(* ================================================================= *)
(*  FB_1030_SafetyManager                                             *)
(*  全机安全管理块: 安全回路状态 + 两次复位 + 启动许可 + 门锁开门流程   *)
(*  版本: V1.0.0  日期: 2026-10-22                                    *)
(*  来源: SysLib/safety/                                              *)
(*  依据: 电气自动化安全规范 V1.0 第 0/2/3/4/5/8/9/12 节               *)
(*        安全FB设计草案_20261022 (用户 10-22 定: 合成一块)            *)
(*  依赖: FB_TON V3.0.0 (真实毫秒), FB_R_TRIG                          *)
(*                                                                    *)
(*  它管什么:                                                         *)
(*    - 只读安全器件报给 PLC 的状态点, 算出"能不能动""复位采不采纳"    *)
(*      "能不能开门", 交给各工位块使用. 全机只调用一次.                *)
(*  它不管什么:                                                       *)
(*    - 不控制安全回路 (回路靠安全继电器硬件切断, 规范 0.1)            *)
(*    - 不决定电磁阀急停后清零还是保持 (工位块按 IO 表, 规范 2.3)       *)
(*    - 不决定断点续跑还是重新初始化 (工位块按项目需求, 规范 2.5)       *)
(*    - 不做光栅屏蔽 (规范 5.3), 不做按钮卡住判断 (规范 3.5)           *)
(*                                                                    *)
(*  状态 q_iState:                                                    *)
(*    0 安全回路断开   1 等满 10 s   2 等运行复位   3 等启动   4 运行许可 *)
(*                                                                    *)
(*  两次复位 (规范 3.1~3.6, 10 s 从第一次按复位起算, 用户 10-21 定):  *)
(*    第一次: 安全继电器自行复位, PLC 只记时刻 (门锁好、总线在线才记)  *)
(*    第二次: 继电器反馈正常 且 距第一次 >= 10 s 才采纳 -> 运行复位脉冲 *)
(*    之后按启动 -> 启动脉冲 + 运行许可. 复位/启动都只认上升沿.         *)
(*                                                                    *)
(*  报警字 q_dwAlarm:                                                 *)
(*    bit0~7   第 1~8 个急停被按下 (实时)                              *)
(*    bit8~15  第 1~8 扇门没关好/没锁 (实时)                           *)
(*    bit16~23 第 1~8 道光栅被遮挡 (实时)                              *)
(*    bit24~27 第 1~4 个安全继电器反馈 = 故障 (实时)                    *)
(*    bit28    总线断线 (实时)                                         *)
(*    bit29    复位被拒: 安全回路未恢复/门没锁/总线断 (保持到下次采纳)  *)
(*    bit30    复位过早: 距第一次不足 10 s (保持到下次采纳)             *)
(*    bit31    门锁回失败: 撤销解锁后 1 s 内门锁点没回来 (保持到锁好)   *)
(*                                                                    *)
(*  安全区: 改本块等于改安全区, 先仿真再由用户签字 (规范 0.5)         *)
(* ================================================================= *)

FUNCTION_BLOCK FB_1030_SafetyManager

VAR_INPUT
    i_arrSafetyFault : ARRAY[0..3] OF BOOL;  // 安全继电器 41-42 常闭辅助点, 1 = 安全回路故障; 未用的填 FALSE (规范 8.1, 判断的唯一依据)
    i_arrEStopOk     : ARRAY[0..7] OF BOOL;  // 急停按钮第三组触点, 1 = 正常; 未用的填 TRUE (规范 2.2, 只报警定位)
    i_arrCurtainOk   : ARRAY[0..7] OF BOOL;  // 光栅进 PLC 的状态点, 1 = 未遮挡; 未用的填 TRUE (规范 5.1, 只报警定位)
    i_arrDoorClosed  : ARRAY[0..7] OF BOOL;  // 门锁进 PLC 的那组触点, 1 = 门关好且已锁; 未用的填 TRUE (规范 4.1, 4.4)
    i_bFieldbusOk    : BOOL;                 // 远程 IO/总线伺服全部在线 (项目汇总后接入, 规范 8.3)
    i_bResetBtn      : BOOL;                 // 复位按钮进 PLC 的那组触点 (规范 3.1)
    i_bStartBtn      : BOOL;                 // 启动按钮 (规范 3.6)
    i_bAutoMode      : BOOL;                 // 设备在自动 (全机一个, 自动时申请开门不响应)
    i_bMotionStopped : BOOL;                 // 伺服零速 + 所有动作完全停止 (全机一个, 项目汇总后接入)
    i_arrDoorReqBtn  : ARRAY[0..7] OF BOOL;  // 每扇门的申请开门按钮; 未用的填 FALSE
END_VAR

VAR_OUTPUT
    q_bSafeToRun     : BOOL;                 // 1 = 可以动; 各工位块的运动输出都要和它"与" (规范 0.1)
    q_bStopNow       : BOOL;                 // 1 = 安全条件现在丢了 (继电器故障/门没锁/总线断), 同一扫描生效 (规范 2.3)
    q_bRunResetPulse : BOOL;                 // 第二次复位被采纳时出一个扫描的脉冲, 清工位故障和握手锁 (规范 3.4)
    q_bStartPulse    : BOOL;                 // 复位以后按启动, 出一个扫描的脉冲 (规范 3.6)
    q_iState         : INT;                  // 状态号 0~4, HMI 显示"现在卡在哪一步"
    q_dwAlarm        : DWORD;                // 报警字, 位定义见文件头
    q_arrDoorUnlock  : ARRAY[0..7] OF BOOL;  // 每扇门的解锁线圈 (得电解锁、失电锁定)
    q_arrDoorLamp    : ARRAY[0..7] OF BOOL;  // 每扇门申请按钮指示灯 (申请中 1 s 周期闪, 允许开门常亮)
END_VAR

VAR
    s_iState         : INT := 0;             // 复位状态机 (上电从 0 开始, 必须人工复位 + 启动)
    s_arrDoorStep    : ARRAY[0..7] OF INT;   // 开门流程 0 锁住 1 申请中 2 允许开门 3 锁回确认
    s_bRejectLatch   : BOOL := FALSE;        // bit29 复位被拒 (保持)
    s_bEarlyLatch    : BOOL := FALSE;        // bit30 复位过早 (保持)
    s_bRelockFail    : BOOL := FALSE;        // bit31 门锁回失败 (保持到所有门锁好)
    s_bDelayRestart  : BOOL := FALSE;        // 本扫描重新开始 10 s 计时 (定时器 IN 断开一拍)
    s_bBlink         : BOOL := FALSE;        // 申请中指示灯闪烁电平

    // ===== 定时器 (先设 IN/PT, 末尾集中调用; FB_TON 真实毫秒) =====
    s_tResetDelay    : FB_TON;               // 第一次复位起的 10 s
    s_tBlink         : FB_TON;               // 闪烁半周期
    s_arrRelockTimer : ARRAY[0..7] OF FB_TON; // 撤销解锁后等门锁点回来

    // ===== 边沿检测 (只认上升沿, 规范 3.1) =====
    s_rtReset        : FB_R_TRIG;
    s_rtStart        : FB_R_TRIG;
    s_arrRtDoorReq   : ARRAY[0..7] OF FB_R_TRIG;
END_VAR

VAR_TEMP
    t_iIdx           : INT;
    t_bFault         : BOOL;                 // 任一安全继电器反馈 = 故障
    t_bDoorsOk       : BOOL;                 // 所有门关好且已锁
    t_bResetEdge     : BOOL;
    t_bStartEdge     : BOOL;
    t_bDelayDone     : BOOL;                 // 距第一次复位已满 10 s (上一扫描定时器结果)
    t_dwBit          : DWORD;
    t_dwAlarm        : DWORD;
END_VAR

VAR CONSTANT
    RESET_DELAY_MS   : DINT := 10000;        // 两次复位最小间隔 10 s (规范 3.4/9, 固定, HMI 不能改)
    BLINK_HALF_MS    : DINT := 500;          // 申请中指示灯 1 s 周期闪烁的半周期 (规范 4.3/9)
    RELOCK_CHECK_MS  : DINT := 1000;         // 撤销解锁后门锁点须在 1 s 内回来, 否则重新解锁 (门开着按复位不采纳)
    ST_OPEN          : INT := 0;             // 安全回路断开
    ST_WAIT_DELAY    : INT := 1;             // 等满 10 s
    ST_WAIT_RESET    : INT := 2;             // 等运行复位
    ST_WAIT_START    : INT := 3;             // 等启动
    ST_RUN           : INT := 4;             // 运行许可
    DOOR_LOCKED      : INT := 0;
    DOOR_REQUEST     : INT := 1;
    DOOR_UNLOCKED    : INT := 2;
    DOOR_RELOCK      : INT := 3;
END_VAR

BEGIN
    (* ================================================================== *)
    (*  1. 读输入: 边沿、汇总                                              *)
    (* ================================================================== *)
    s_rtReset(IN := i_bResetBtn);
    t_bResetEdge := s_rtReset.Q;
    s_rtStart(IN := i_bStartBtn);
    t_bStartEdge := s_rtStart.Q;
    t_bDelayDone := s_tResetDelay.Q;

    t_bFault := FALSE;
    FOR t_iIdx := 0 TO 3 DO
        t_bFault := t_bFault OR i_arrSafetyFault[t_iIdx];
    END_FOR;
    t_bDoorsOk := TRUE;
    FOR t_iIdx := 0 TO 7 DO
        t_bDoorsOk := t_bDoorsOk AND i_arrDoorClosed[t_iIdx];
    END_FOR;

    q_bRunResetPulse := FALSE;
    q_bStartPulse := FALSE;
    s_bDelayRestart := FALSE;

    (* ================================================================== *)
    (*  2. 任何状态: 继电器故障/门没锁/总线断 -> 当拍回状态 0             *)
    (*     状态 1 在等继电器自己复位, 继电器故障是预期的, 只看门和总线      *)
    (* ================================================================== *)
    IF s_iState >= ST_WAIT_RESET THEN
        IF t_bFault OR NOT t_bDoorsOk OR NOT i_bFieldbusOk THEN
            s_iState := ST_OPEN;
        END_IF;
    ELSIF s_iState = ST_WAIT_DELAY THEN
        IF NOT t_bDoorsOk OR NOT i_bFieldbusOk THEN
            s_iState := ST_OPEN;
        END_IF;
    END_IF;

    (* ================================================================== *)
    (*  3. 两次复位状态机 (规范第 3 节)                                     *)
    (* ================================================================== *)
    CASE s_iState OF
        ST_OPEN:
            // 第一次复位: 只记时刻, 不清任何东西. 门没锁或总线断时继电器也复位不了, 不记, 报复位被拒
            IF t_bResetEdge THEN
                IF t_bDoorsOk AND i_bFieldbusOk THEN
                    s_bRejectLatch := FALSE;
                    s_bEarlyLatch := FALSE;
                    s_bDelayRestart := TRUE;
                    s_iState := ST_WAIT_DELAY;
                ELSE
                    s_bRejectLatch := TRUE;
                END_IF;
            END_IF;

        ST_WAIT_DELAY:
            IF t_bDelayDone AND NOT t_bFault THEN
                // 满 10 s 且反馈正常: 可以按第二次了
                s_iState := ST_WAIT_RESET;
            ELSIF t_bResetEdge THEN
                IF t_bDelayDone THEN
                    // 10 s 到了反馈仍不正常, 这一下当作新的第一次, 重新计 10 s
                    s_bRejectLatch := FALSE;
                    s_bEarlyLatch := FALSE;
                    s_bDelayRestart := TRUE;
                ELSIF t_bFault THEN
                    s_bRejectLatch := TRUE;   // 安全回路未恢复, 不采纳
                ELSE
                    s_bEarlyLatch := TRUE;    // 不足 10 s, 不采纳
                END_IF;
            ELSIF t_bDelayDone AND t_bFault THEN
                s_bRejectLatch := TRUE;       // 10 s 到了安全回路仍未恢复, 等重新按第一次
            END_IF;

        ST_WAIT_RESET:
            // 第二次复位: 反馈正常、门锁好、总线在线已由第 2 段保证
            IF t_bResetEdge THEN
                q_bRunResetPulse := TRUE;
                s_bRejectLatch := FALSE;
                s_bEarlyLatch := FALSE;
                s_iState := ST_WAIT_START;
            END_IF;

        ST_WAIT_START:
            IF t_bStartEdge THEN
                q_bStartPulse := TRUE;
                s_iState := ST_RUN;
            ELSIF t_bResetEdge THEN
                // 已复位还没启动时按复位: 只清报警, 不出脉冲
                s_bRejectLatch := FALSE;
                s_bEarlyLatch := FALSE;
            END_IF;

        ST_RUN:
            // 运行许可: 只有第 2 段 (安全条件丢失) 能让它离开
            s_bDelayRestart := FALSE;

        ELSE
            s_iState := ST_OPEN;
    END_CASE;

    (* ================================================================== *)
    (*  4. 开门流程 (规范 4.3): 每扇门一套, 下标 0~7 = 第 1~8 扇门         *)
    (* ================================================================== *)
    FOR t_iIdx := 0 TO 7 DO
        s_arrRtDoorReq[t_iIdx](IN := i_arrDoorReqBtn[t_iIdx]);

        CASE s_arrDoorStep[t_iIdx] OF
            DOOR_LOCKED:
                // 自动时按申请不响应
                IF s_arrRtDoorReq[t_iIdx].Q AND NOT i_bAutoMode THEN
                    s_arrDoorStep[t_iIdx] := DOOR_REQUEST;
                END_IF;

            DOOR_REQUEST:
                IF i_bAutoMode THEN
                    s_arrDoorStep[t_iIdx] := DOOR_LOCKED;      // 申请中切回自动, 取消申请
                ELSIF i_bMotionStopped THEN
                    s_arrDoorStep[t_iIdx] := DOOR_UNLOCKED;    // 伺服停、动作全停, 允许开门
                END_IF;

            DOOR_UNLOCKED:
                // 关门后按复位: 撤销解锁, 去确认门锁点回来
                IF t_bResetEdge THEN
                    s_arrDoorStep[t_iIdx] := DOOR_RELOCK;
                END_IF;

            DOOR_RELOCK:
                IF i_arrDoorClosed[t_iIdx] THEN
                    s_arrDoorStep[t_iIdx] := DOOR_LOCKED;
                ELSIF s_arrRelockTimer[t_iIdx].Q THEN
                    // 1 s 内门锁点没回来 = 门还开着, 这次复位不采纳, 恢复解锁 (人可能还在里面)
                    s_bRelockFail := TRUE;
                    s_arrDoorStep[t_iIdx] := DOOR_UNLOCKED;
                END_IF;

            ELSE
                s_arrDoorStep[t_iIdx] := DOOR_LOCKED;
        END_CASE;

        s_arrRelockTimer[t_iIdx].IN := (s_arrDoorStep[t_iIdx] = DOOR_RELOCK);
        s_arrRelockTimer[t_iIdx].PT := RELOCK_CHECK_MS;
    END_FOR;
    IF t_bDoorsOk THEN
        s_bRelockFail := FALSE;
    END_IF;

    // 申请中指示灯 1 s 周期闪烁: 半周期定时器自复位, 到时翻转
    s_tBlink.IN := NOT s_tBlink.Q;
    s_tBlink.PT := BLINK_HALF_MS;
    IF s_tBlink.Q THEN
        s_bBlink := NOT s_bBlink;
    END_IF;

    FOR t_iIdx := 0 TO 7 DO
        q_arrDoorUnlock[t_iIdx] := (s_arrDoorStep[t_iIdx] = DOOR_UNLOCKED);
        q_arrDoorLamp[t_iIdx] := (s_arrDoorStep[t_iIdx] = DOOR_UNLOCKED)
                                 OR ((s_arrDoorStep[t_iIdx] = DOOR_REQUEST) AND s_bBlink);
    END_FOR;

    (* ================================================================== *)
    (*  5. 定时器集中调用                                                  *)
    (* ================================================================== *)
    s_tResetDelay.IN := (s_iState = ST_WAIT_DELAY) AND NOT s_bDelayRestart;
    s_tResetDelay.PT := RESET_DELAY_MS;
    s_tResetDelay(IN := s_tResetDelay.IN, PT := s_tResetDelay.PT);
    s_tBlink(IN := s_tBlink.IN, PT := s_tBlink.PT);
    FOR t_iIdx := 0 TO 7 DO
        s_arrRelockTimer[t_iIdx](IN := s_arrRelockTimer[t_iIdx].IN, PT := s_arrRelockTimer[t_iIdx].PT);
    END_FOR;

    (* ================================================================== *)
    (*  6. 输出                                                            *)
    (* ================================================================== *)
    q_iState := s_iState;
    q_bSafeToRun := (s_iState = ST_RUN);
    q_bStopNow := t_bFault OR NOT t_bDoorsOk OR NOT i_bFieldbusOk;

    t_dwAlarm := 16#00000000;
    t_dwBit := 16#00000001;
    FOR t_iIdx := 0 TO 7 DO
        IF NOT i_arrEStopOk[t_iIdx] THEN
            t_dwAlarm := t_dwAlarm OR SHL(t_dwBit, INT_TO_UINT(t_iIdx));
        END_IF;
        IF NOT i_arrDoorClosed[t_iIdx] THEN
            t_dwAlarm := t_dwAlarm OR SHL(t_dwBit, INT_TO_UINT(t_iIdx + 8));
        END_IF;
        IF NOT i_arrCurtainOk[t_iIdx] THEN
            t_dwAlarm := t_dwAlarm OR SHL(t_dwBit, INT_TO_UINT(t_iIdx + 16));
        END_IF;
    END_FOR;
    FOR t_iIdx := 0 TO 3 DO
        IF i_arrSafetyFault[t_iIdx] THEN
            t_dwAlarm := t_dwAlarm OR SHL(t_dwBit, INT_TO_UINT(t_iIdx + 24));
        END_IF;
    END_FOR;
    IF NOT i_bFieldbusOk THEN
        t_dwAlarm := t_dwAlarm OR SHL(t_dwBit, 28);
    END_IF;
    IF s_bRejectLatch THEN
        t_dwAlarm := t_dwAlarm OR SHL(t_dwBit, 29);
    END_IF;
    IF s_bEarlyLatch THEN
        t_dwAlarm := t_dwAlarm OR SHL(t_dwBit, 30);
    END_IF;
    IF s_bRelockFail THEN
        t_dwAlarm := t_dwAlarm OR SHL(t_dwBit, 31);
    END_IF;
    q_dwAlarm := t_dwAlarm;

END_FUNCTION_BLOCK
